FUNCTION_BLOCK AOption_AUI_DEMUX_1 (* AOption demultiplexor (generic FB): aktiviert per Index K genau einen von 1 Options-Ausgaengen (INIT_REQ), kein IN-Wert noetig. *)
  (* Standard: 61499-2; Description: Copyright (c) 2026 Meisterschulen am Ostbahnhof This program and the accompanying materials are made available under the terms of the Eclipse Public License 2.0 which is available at https://www.eclipse.org/legal/epl-2.0/ SPDX-License-Identifier: EPL-2.0 *)
  (* Version 1.0, 2026-10-13, Franz Höpfinger, Meisterschulen am Ostbahnhof *)
  PACKAGE Option::selection;
  {SET_ATTRIBUTE(eclipse4diac::core::GenericClassName, 'GEN_AOption_AUI_DEMUX')}
  (* Documentation:
  Demultiplexer (natives Generic-FB, kein ECC/Algorithmus in diesem Typ) fuer N=1 Options-Ausgaenge vom Typ Option::AOption, ausgewaehlt ueber den bidirektionalen Index-Adapter K (adapter::types::bidirectional::AUI2).
   Indexzuordnung:
    - K = 0 – alle Ausgaenge AUS
   - K = 1 – OUT1 AN, alle anderen AUS
   - jeder andere Wert (negativ, > 1, ...) – alle Ausgaenge AUS
    Umschaltverhalten (Break-before-Make): wechselt K z.B. von 1 auf 2, wird zuerst der bisher aktive Ausgang (OUT1) deaktiviert (INIT_REQ mit QI=FALSE). Erst wenn von diesem Ausgang die Bestaetigung INIT_CNF eingetroffen ist, wird der neu ausgewaehlte Ausgang (OUT2) aktiviert (INIT_REQ mit QI=TRUE). Es ist also niemals mehr als eine Option gleichzeitig aktiv.
   Pro eintreffendem K-Wert wird jeder Ausgang maximal 1x getriggert (der zuvor aktive einmal zum Abschalten, der neu ausgewaehlte einmal zum Einschalten) - nicht betroffene Ausgaenge werden nicht angefasst.
   Busy-Gating ueber den bidirektionalen K-Adapter: Waehrend ein Umschaltvorgang laeuft (also solange auf INIT_CNF vom bisherigen und/oder neuen Ausgang gewartet wird), wird jeder weitere ueber K (Richtung Plug -> Socket, EO1/DO1) eintreffende Indexwunsch ignoriert - er wird weder gepuffert noch nachgeholt. Erst wenn der Umschaltvorgang abgeschlossen ist, meldet der DEMUX dies rueckwaerts ueber K (Richtung Socket -> Plug, EI1/DI1) mit dem uebernommenen K-Wert zurueck (nicht mit dem Zustand der Ausgaenge: auch ein ungueltiger Wert wird unveraendert quittiert); erst danach werden wieder neue Indexwuensche angenommen. Damit sind sowohl langsame Umschaltvorgaenge (lange Reaktionszeit der Ausgaenge) als auch mehrfache, einander widersprechende K-Werte in kurzer Folge sauber abgedeckt: es zaehlt immer nur der Stand nach Abschluss des letzten tatsaechlich bearbeiteten Wechsels.
  *)
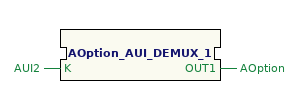
  SOCKETS
    K : adapter::types::bidirectional::AUI2; (* index (bidirektional: EO1/DO1 = neuer K-Wunsch rein, EI1/DI1 = Quittung mit dem uebernommenen Wert zurueck) *)
  END_SOCKETS
  PLUGS
    OUT1 : Option::AOption; (* Option 1 (ausgewaehlt wenn K = 1) *)
  END_PLUGS
END_FUNCTION_BLOCK
